// TIA Portal V19 export
TYPE "ST_Servo"
   STRUCT
      Move : "ST_Move";
      Home : "ST_Home";
      Power : "ST_Power";
      Reset : "ST_Reset";
      Jogging : "ST_Joggong";
   END_STRUCT;
END_TYPE
